(* IEC 61131-3 sources: BODAS-RC27-18_40/st/bodas_rc18_12_27_18_40/plc_logic/application/easyconfig_import/bds_sent_ec, 2 files *)

(* ---- bds_sent_signal_te-bds_sent_signal_te.st ---- *)
(* --- Interface --- *)
///Definition configuration of available SENT signals (consists signals of all variants)
{attribute 'qualified_only' := ''}
{attribute 'strict' := ''}
TYPE bds_sent_signal_te :
(
	///X_X_X04
	bds_sent_K59_E := 0,
	///X_X_X19
	bds_sent_K56_E,
	bds_sent_numSignal_E
) USINT;
END_TYPE

(* ---- bds_sent_ec_gvl-bds_sent_ec_gvl.st ---- *)
(* --- Interface --- *)
{attribute 'qualified_only' := ''}
VAR_GLOBAL CONSTANT
	bds_sent_postVariants_du8: USINT := 1;
	bds_sent_maxDataNibbles_du8: USINT := 6;
	bds_sent_rxFastDataBufSize_du8: USINT := 0;
	bds_sent_rxSlowDataBufSize_du8: USINT := 0;
END_VAR
